// TIA Portal V20 export
VAR_GLOBAL   // PLC tag table "memor"
   HSC_1 AT %ID1000 : DWord;
   PAMET_TEST AT %MD16 : DInt;
   ret_val_move_blk AT %MW20 : Int;
   i AT %MW22 : Int;
   "i(1)" AT %MW24 : Int;
END_VAR
